{attribute 'analysis' := '-33'}
PROGRAM PRG_TEST
VAR
    (* Seeds PMPS_GVL.BP_jsonDoc with the fake test PMPS DB in before any test FB body runs. *)
    fbPmpsTestSetup: FB_CC_PMPSTestSetup;
    fbATMTest: FB_ATMTest;
    fbGBSTest: FB_GBSTest;
    fbIPMTest: FB_IPMTest;
    fbLICTest: FB_LICTest;
    fbPPMTest: FB_PPMTest;
    fbREFTest: FB_REFTest;
    fbSATTTest: FB_SATTTest;
    fbSlitsPowerTest: FB_SLITS_POWERTest;
    fbWFSTest: FB_WFSTest;
    fbXPIMTest: FB_XPIMTest;
    fbCCTempSensorTest: FB_CC_TempSensorTest;


END_VAR

// Run the tests
TcUnit.RUN();

END_PROGRAM

(* stored: Version 1.1.0.1
   POU PRG_TEST: Id {f53165b1-b00c-43dc-a7bd-df3f4a7d5ece}, SpecialFunc None *)
